Fanuc KAREL source: kd00051.KL

-- PROVISIONAL review KL for V770-1; original PC SHA256 92656b6c98507c3d1e9eba6e170f882512f6b5617ebfe71904c4de4527f7f1f1
-- Incomplete behavior may be omitted. Consult companion uncertainty JSON. Do not deploy.
PROGRAM KD00051
%NOLOCKGROUP
VAR
  I : INTEGER
  J : INTEGER
  B : BOOLEAN
  R : REAL
  S : STRING[80]
-- UNRESOLVED_DECL P type=000101
BEGIN
  -- UNRESOLVED_PC offsets 5-30; opcodes 01,22,1C,2E,0A,82,0B
  -- UNRESOLVED_PC offsets 35-39; opcodes 7F
END KD00051
